# EPICS substitutions: xrmIocApp/Db/permit_lut_16R.substitutions
file "permit_lut.template"
{
    pattern {ROW0, ADDR}
        {01, 0}
        {02, 1}
        {03, 2}
        {04, 3}
        {05, 4}
        {06, 5}
        {07, 6}
        {08, 7}
        {09, 8}
        {10, 9}
        {11,10}
        {12,11}
        {13,12}
        {14,13}
        {15,14}
        {16,15}
}
